Fanuc KAREL source: KT00531.KL

PROGRAM KT00531
%NOLOCKGROUP
VAR
  P1: XYZWPREXT
  P2: JOINTPOS
  OUT: XYZWPREXT
BEGIN
  P1.X = 1.0
  OUT = P1 : P2
END KT00531
